(*
SPDX-FileCopyrightText: © 2026 Oleksandr Tiutyk <trofimich@gmail.com>
SPDX-License-Identifier: MIT
License: https://opensource.org/license/mit
*)

(*!
<summary>Orders LTIME values described by generic descriptors.</summary>
<description>
Non-null addresses must reference live LTIME storage. TypeClass and Size are not validated and no numeric
conversion is performed. Two null addresses compare equal; one null address sorts before a non-null address.
Descriptors are passed by value; payload remains borrowed and is not modified, cloned, released or retained.
IsMemoryOwner does not affect comparison.
</description>
*)

FUNCTION_BLOCK LTimeComparer EXTENDS TOF_Core.Object IMPLEMENTS TOF_Core.IComparer
VAR_STAT
	//! <summary>Class name shared by all instances of this function block.</summary>
	{attribute 'hide'} 
	_ClassName : STRING := __POUNAME();
END_VAR

{attribute 'monitoring' := 'call'}
PROPERTY ClassName : REFERENCE TO STRING
GET
ClassName REF= _ClassName;
END_GET
END_PROPERTY

(*!
<summary>Compares the first operand with the second using this ordering strategy.</summary>
<description>
Non-null addresses must reference live LTIME storage. TypeClass and Size are not validated and no numeric
conversion is performed. Two null addresses compare equal; one null address sorts before a non-null address.
Descriptors are passed by value; payload remains borrowed and is not modified, cloned, released or retained.
IsMemoryOwner does not affect comparison. Descendants cannot replace this standard ordering; implement
IComparer separately for a different ordering strategy.
</description>
*)
//!<param name="first">First descriptor; referenced storage is borrowed for the call.</param>
//!<param name="second">Second descriptor; referenced storage is borrowed for the call.</param>
{attribute "object_name" := "Compare"}
METHOD FINAL Compare : TOF_Core.COMPARISON_RESULT
VAR_INPUT
	first : TOF_Core.GENERIC_VALUE;
	second : TOF_Core.GENERIC_VALUE;
END_VAR
VAR
	leftPointer : POINTER TO LTIME; 
	rightPointer : POINTER TO LTIME; 
END_VAR
IF first.Address = 0 AND_THEN second.Address = 0 THEN
	Compare := TOF_Core.COMPARISON_RESULT.FIRST_EQUAL_TO_SECOND;
	RETURN;
END_IF

IF first.Address = 0 THEN
	Compare := TOF_Core.COMPARISON_RESULT.FIRST_LESS_THAN_SECOND;
	RETURN;	
END_IF

IF second.Address = 0 THEN
	Compare := TOF_Core.COMPARISON_RESULT.FIRST_GREATER_THAN_SECOND;
	RETURN;	
END_IF

leftPointer := first.Address;
rightPointer := second.Address;

IF leftPointer^ < rightPointer^ THEN
	Compare := TOF_Core.COMPARISON_RESULT.FIRST_LESS_THAN_SECOND;
ELSIF leftPointer^ > rightPointer^ THEN
	Compare := TOF_Core.COMPARISON_RESULT.FIRST_GREATER_THAN_SECOND;
ELSE
	Compare := TOF_Core.COMPARISON_RESULT.FIRST_EQUAL_TO_SECOND;	
END_IF
END_METHOD

{attribute 'monitoring' := 'call'}
PROPERTY NamespaceName : REFERENCE TO STRING
GET
NamespaceName REF= CurrentNamespace.Name;
END_GET
END_PROPERTY

{attribute 'monitoring' := 'call'}
PROPERTY SelfSize : ULINT
GET
SelfSize := XSIZEOF(THIS^);
END_GET
END_PROPERTY

END_FUNCTION_BLOCK

(* stored: Version 1.1.0.1
   POU LTimeComparer: Id {ace72394-daf6-4b9d-a33d-9a436c0a305e}, SpecialFunc None
   Property ClassName: Id {85665c3e-8f5e-44c8-b281-b80838358c8a}
   Get Get: Id {efcaf5c8-16fb-4602-8bb0-efa67641ae20}
   Method Compare: Id {b669a8e2-61ab-4523-b98f-4dc19e868351}
   Property NamespaceName: Id {914a33de-ef85-46ea-a5f0-4f046b7f90db}
   Get Get: Id {e459264c-369a-41e0-bede-f57b12c3f5cb}
   Property SelfSize: Id {589d987c-a708-4ea5-8f21-736c80a729d0}
   Get Get: Id {02fdeab4-5b77-4079-8ffc-c9e19327056c} *)
